(* Logix 5000 project; controller TFF vendor 1 type 14 code 107 rev 33.11; software revision 33.04; part 15 of 38 *)
(* tags used below, declared in another part *)
   ActionCode : DINT;   // Action Code
   AutoRunTimer : TIMER;   // Auto Run Timer
   Clear : BOOL;   // Clear Operation Table Flag
   Criteria1Code : DINT;   // Criteria 1 Code
   Criteria2Code : DINT;   // Criteria 2 Code
   CriteriaMet : BOOL;   // Criteria Met
   DownloadONS : BOOL;
   ErrorCheck : BOOL;   // Error Check Flag
   PhaseClear : BOOL;   // Phase Clear
   PhaseNumber : DINT;   // Phase FOR NEXT Index
   PreRunLog : BOOL;   // Log Pre Run Set Points
   Run : BOOL;   // Operation Run Status
   RunONS : BOOL;   // Run Command One-Shot
   Structure : DINT;   // Structure code
   Value : REAL;   // Temp Value
   AlarmControl : AlarmControl;   // Alarm Control
   CCPSystem : CCPSystem;   // CCP System Data
   CPU_Scanning : BOOL;   // System Scanning Flag
   Memory_Data : Memory_Data;
   Memory_Message : MESSAGE;   // Data for Message instruction read Memory informations
   Memory_Temp : INT[29];   // Destination elements for message read Memory informations
   Operation : Operation[6,251];   // Operation Table
   PCDateTime : DINT[7];   // Date/Time Array from PC
   Phase : Phases[6];   // Phase Control Array
   Phase0 : ALIAS FOR Phase[0];   // Phase 0
   PLCFault : FaultRecordType;   // PLC Major Fault Record
   Prompt : Prompt[7];   // Prompt Array
   Prompt0 : ALIAS FOR Prompt[0];   // Phase 0 Prompt
   Prompt1 : ALIAS FOR Prompt[1];   // Phase 1 Prompt
   Prompt2 : ALIAS FOR Prompt[2];   // Phase 2 Prompt
   Prompt3 : ALIAS FOR Prompt[3];   // Phase 3 Prompt
   Prompt4 : ALIAS FOR Prompt[4];   // Phase 4 Prompt
   Prompt5 : ALIAS FOR Prompt[5];   // Phase 5 Prompt
   ResumeDownloadFromHOLD : BOOL;   // Resume Download From HOLD
   TimerControl : TimerControl;   // Timer Control
   Timers : Timers[22];   // Timer Array
   YA10 : ALIAS FOR DigitalPoint[59];
(* CCPSystem, continued *)

ROUTINE Prompt   (* ladder *)
// Operator Prompt Routine
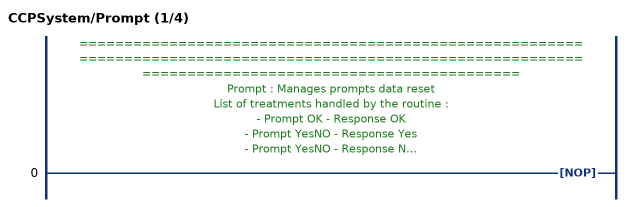
   // ==========================================================================================================================================================
   //                                                                                                                       Prompt : Manages prompts data reset
   //                                                     List of treatments handled by the routine :
   //                                                          - Prompt OK - Response OK
   //                                                          - Prompt YesNO - Response Yes
   //                                                          - Prompt YesNO - Response No
   //                                                     -----------------------------------------------------------------------------------------------------------------------------------------------------
   //                                                     History
   // 		2019-DEC-24 - Merck - Q. Spindler - Initial version for Candidate Release 1.00.00.00.a
   // 		2022-SEP-20 - Actemium - J. Jaekel - Modification for Candidate Release 1.01.00.01.a
   // - Add condition to avoid discarding the prompt response on other phases than 0
   // ============================================================================================================================
   // ============================
   0: NOP();
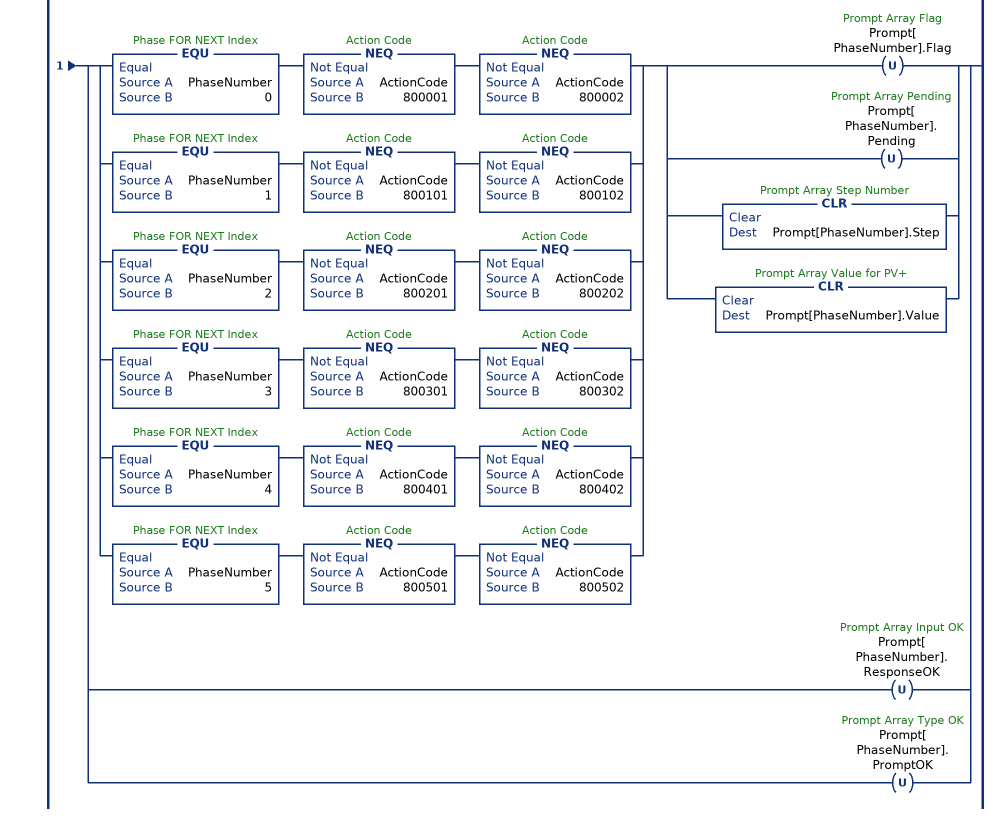
   // Prompt OK - Response OK
   // ==========================================================================================================================================================
   1: XIC(Prompt[PhaseNumber].PromptOK)XIC(Prompt[PhaseNumber].ResponseOK)[XIC(CriteriaMet) ,XIC(Phase[PhaseNumber].JumpPLC) ,EQU(PhaseNumber,0) NEQ(Criteria1Code,800003) NEQ(Criteria2Code,800003) ,EQU(PhaseNumber,1) NEQ(Criteria1Code,800103) NEQ(Criteria2Code,800103) ,EQU(PhaseNumber,2) NEQ(Criteria1Code,800203) NEQ(Criteria2Code,800203) ,EQU(PhaseNumber,3) NEQ(Criteria1Code,800303) NEQ(Criteria2Code,800303) ,EQU(PhaseNumber,4) NEQ(Criteria1Code,800403) NEQ(Criteria2Code,800403) ,EQU(PhaseNumber,5) NEQ(Criteria1Code,800503) NEQ(Criteria2Code,800503) ][[EQU(PhaseNumber,0) NEQ(ActionCode,800001) NEQ(ActionCode,800002) ,EQU(PhaseNumber,1) NEQ(ActionCode,800101) NEQ(ActionCode,800102) ,EQU(PhaseNumber,2) NEQ(ActionCode,800201) NEQ(ActionCode,800202) ,EQU(PhaseNumber,3) NEQ(ActionCode,800301) NEQ(ActionCode,800302) ,EQU(PhaseNumber,4) NEQ(ActionCode,800401) NEQ(ActionCode,800402) ,EQU(PhaseNumber,5) NEQ(ActionCode,800501) NEQ(ActionCode,800502) ] [OTU(Prompt[PhaseNumber].Flag) ,OTU(Prompt[PhaseNumber].Pending) ,CLR(Prompt[PhaseNumber].Step) ,CLR(Prompt[PhaseNumber].Value) ] ,OTU(Prompt[PhaseNumber].ResponseOK) ,OTU(Prompt[PhaseNumber].PromptOK) ];
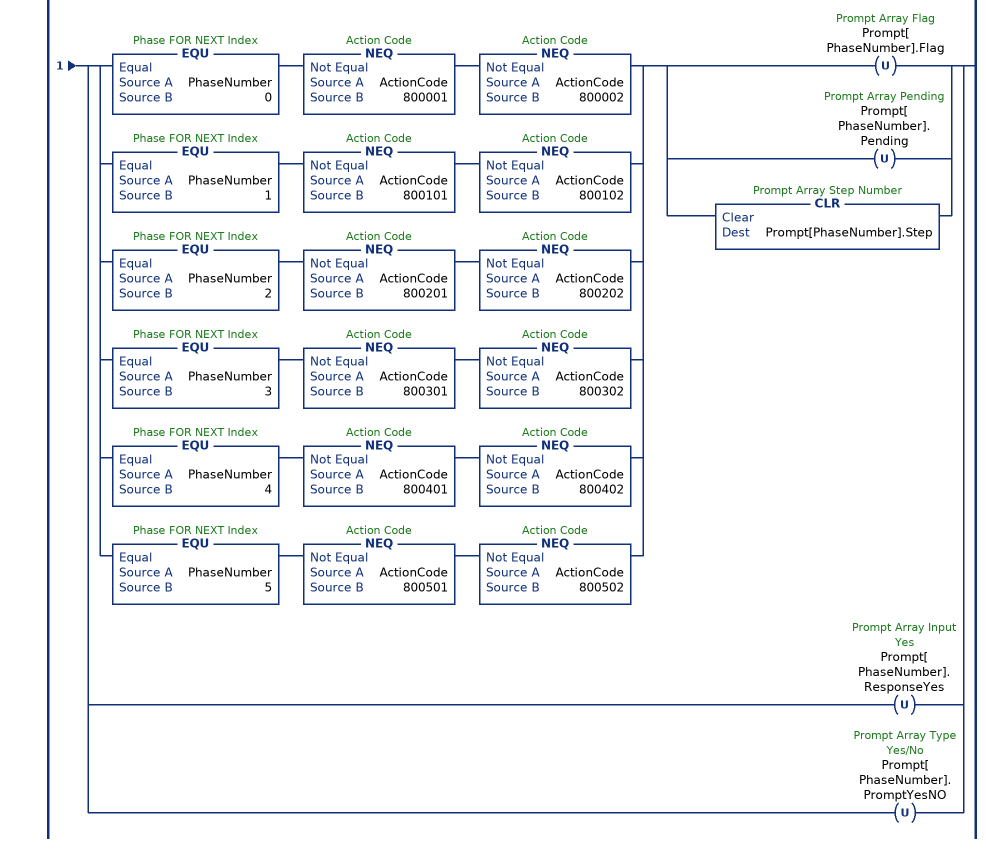
   // Prompt YesNO - Response Yes
   // ==========================================================================================================================================================
   2: XIC(Prompt[PhaseNumber].PromptYesNO)XIC(Prompt[PhaseNumber].ResponseYes)[XIC(CriteriaMet) ,XIC(Phase[PhaseNumber].JumpPLC) ,EQU(PhaseNumber,0) NEQ(Criteria1Code,800004) NEQ(Criteria2Code,800004) ,EQU(PhaseNumber,1) NEQ(Criteria1Code,800104) NEQ(Criteria2Code,800104) ,EQU(PhaseNumber,2) NEQ(Criteria1Code,800204) NEQ(Criteria2Code,800204) ,EQU(PhaseNumber,3) NEQ(Criteria1Code,800304) NEQ(Criteria2Code,800304) ,EQU(PhaseNumber,4) NEQ(Criteria1Code,800404) NEQ(Criteria2Code,800404) ,EQU(PhaseNumber,5) NEQ(Criteria1Code,800504) NEQ(Criteria2Code,800504) ][[EQU(PhaseNumber,0) NEQ(ActionCode,800001) NEQ(ActionCode,800002) ,EQU(PhaseNumber,1) NEQ(ActionCode,800101) NEQ(ActionCode,800102) ,EQU(PhaseNumber,2) NEQ(ActionCode,800201) NEQ(ActionCode,800202) ,EQU(PhaseNumber,3) NEQ(ActionCode,800301) NEQ(ActionCode,800302) ,EQU(PhaseNumber,4) NEQ(ActionCode,800401) NEQ(ActionCode,800402) ,EQU(PhaseNumber,5) NEQ(ActionCode,800501) NEQ(ActionCode,800502) ] [OTU(Prompt[PhaseNumber].Flag) ,OTU(Prompt[PhaseNumber].Pending) ,CLR(Prompt[PhaseNumber].Step) ] ,OTU(Prompt[PhaseNumber].ResponseYes) ,OTU(Prompt[PhaseNumber].PromptYesNO) ];
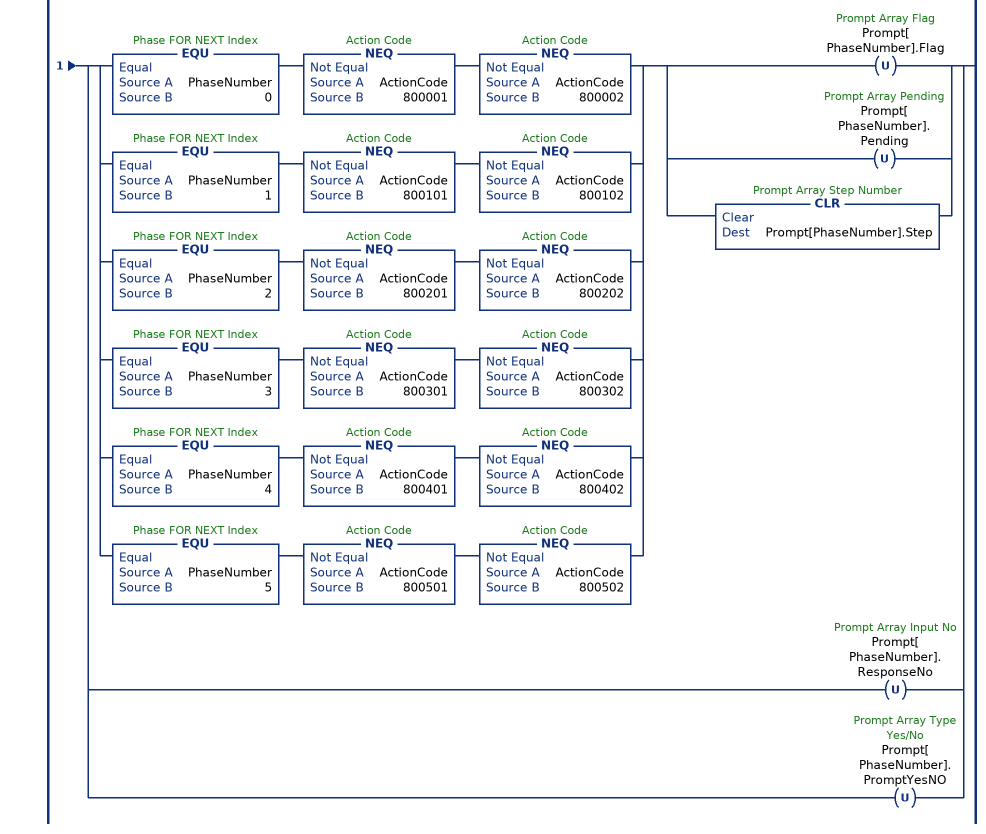
   // Prompt YesNO - Response No
   // ==========================================================================================================================================================
   3: XIC(Prompt[PhaseNumber].PromptYesNO)XIC(Prompt[PhaseNumber].ResponseNo)[XIC(CriteriaMet) ,XIC(Phase[PhaseNumber].JumpPLC) ,EQU(PhaseNumber,0) NEQ(Criteria1Code,800005) NEQ(Criteria2Code,800005) ,EQU(PhaseNumber,1) NEQ(Criteria1Code,800105) NEQ(Criteria2Code,800105) ,EQU(PhaseNumber,2) NEQ(Criteria1Code,800205) NEQ(Criteria2Code,800205) ,EQU(PhaseNumber,3) NEQ(Criteria1Code,800305) NEQ(Criteria2Code,800305) ,EQU(PhaseNumber,4) NEQ(Criteria1Code,800405) NEQ(Criteria2Code,800405) ,EQU(PhaseNumber,5) NEQ(Criteria1Code,800505) NEQ(Criteria2Code,800505) ][[EQU(PhaseNumber,0) NEQ(ActionCode,800001) NEQ(ActionCode,800002) ,EQU(PhaseNumber,1) NEQ(ActionCode,800101) NEQ(ActionCode,800102) ,EQU(PhaseNumber,2) NEQ(ActionCode,800201) NEQ(ActionCode,800202) ,EQU(PhaseNumber,3) NEQ(ActionCode,800301) NEQ(ActionCode,800302) ,EQU(PhaseNumber,4) NEQ(ActionCode,800401) NEQ(ActionCode,800402) ,EQU(PhaseNumber,5) NEQ(ActionCode,800501) NEQ(ActionCode,800502) ] [OTU(Prompt[PhaseNumber].Flag) ,OTU(Prompt[PhaseNumber].Pending) ,CLR(Prompt[PhaseNumber].Step) ] ,OTU(Prompt[PhaseNumber].ResponseNo) ,OTU(Prompt[PhaseNumber].PromptYesNO) ];
END_ROUTINE

ROUTINE Start   (* ladder *)
// Operation Start Routine
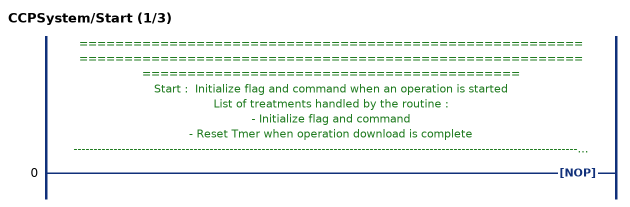
   // ==========================================================================================================================================================
   //                                                                                                      Start :  Initialize flag and command when an operation is started
   //                                                     List of treatments handled by the routine :
   //                                                          - Initialize flag and command
   //                                                          - Reset Tmer when operation download is complete
   //                                                     -----------------------------------------------------------------------------------------------------------------------------------------------------
   //                                                     History
   // 		2019-DEC-24 - Merck - Q. Spindler - Initial version for Candidate Release 1.00.00.00.a
   // ========================================================================================================================================================
   0: NOP();
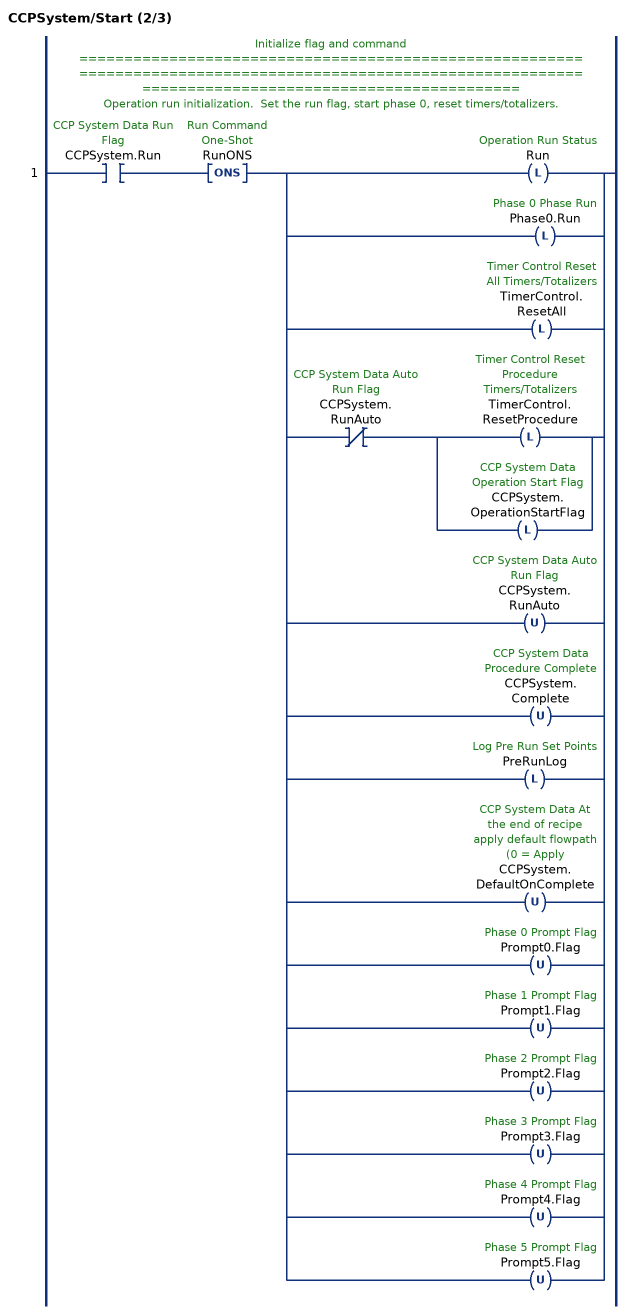
   // Initialize flag and command
   // ==========================================================================================================================================================
   // Operation run initialization.  Set the run flag, start phase 0, reset timers/totalizers.
   1: XIC(CCPSystem.Run)ONS(RunONS)[OTL(Run) ,OTL(Phase0.Run) ,OTL(TimerControl.ResetAll) ,XIO(CCPSystem.RunAuto) [OTL(TimerControl.ResetProcedure) ,OTL(CCPSystem.OperationStartFlag) ] ,OTU(CCPSystem.RunAuto) ,OTU(CCPSystem.Complete) ,OTL(PreRunLog) ,OTU(CCPSystem.DefaultOnComplete) ,OTU(Prompt0.Flag) ,OTU(Prompt1.Flag) ,OTU(Prompt2.Flag) ,OTU(Prompt3.Flag) ,OTU(Prompt4.Flag) ,OTU(Prompt5.Flag) ];
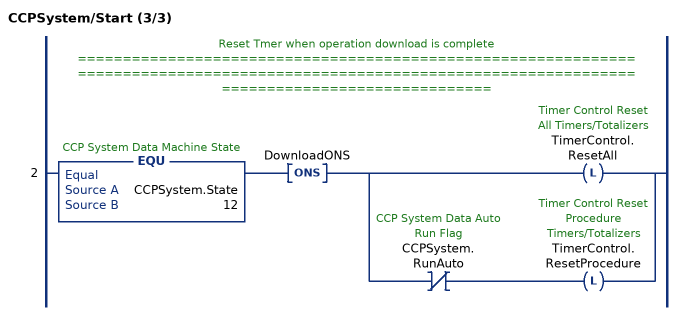
   // Reset Tmer when operation download is complete
   // ==========================================================================================================================================================
   2: EQU(CCPSystem.State,12)ONS(DownloadONS)[OTL(TimerControl.ResetAll) ,XIO(CCPSystem.RunAuto) OTL(TimerControl.ResetProcedure) ];
END_ROUTINE

ROUTINE State   (* ladder *)
// Machine State Routine
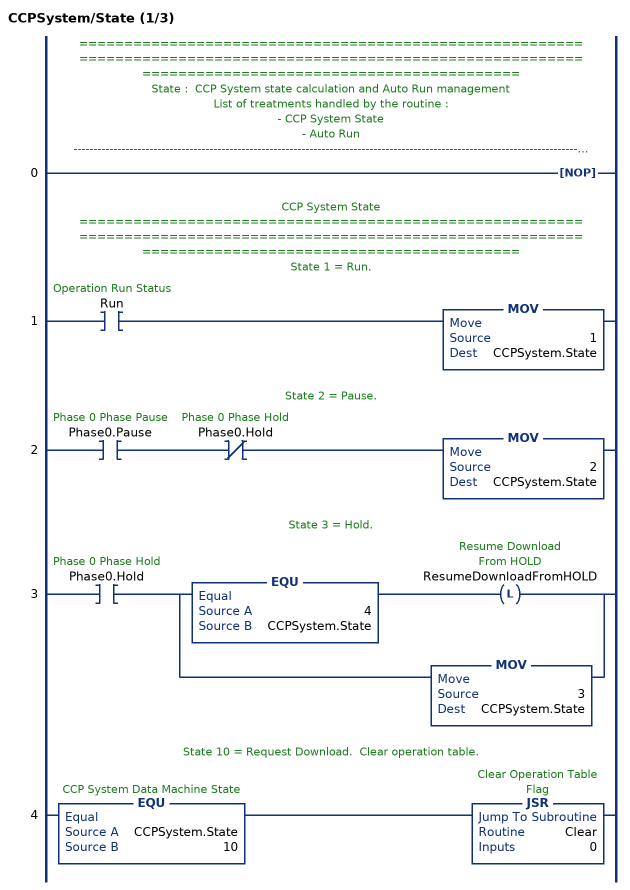
   // ==========================================================================================================================================================
   //                                                                                                  State :  CCP System state calculation and Auto Run management
   //                                                     List of treatments handled by the routine :
   //                                                          - CCP System State
   //                                                          - Auto Run
   //                                                     -----------------------------------------------------------------------------------------------------------------------------------------------------
   //                                                     History
   // 		2019-DEC-24 - Merck - Q. Spindler - Initial version for Candidate Release 1.00.00.00.a
   // 		2021-APR-22 - Merck - Q. Spindler - Modifications for Candidate Release 1.00.00.00.e
   // - Add of Resume Download From HOLD state
   // ========================================================================================================================================================
   0: NOP();
   // CCP System State
   // ==========================================================================================================================================================
   // State 1 = Run.
   1: XIC(Run)MOV(1,CCPSystem.State);
   // State 2 = Pause.
   2: XIC(Phase0.Pause)XIO(Phase0.Hold)MOV(2,CCPSystem.State);
   // State 3 = Hold.
   3: XIC(Phase0.Hold)[EQU(4,CCPSystem.State) OTL(ResumeDownloadFromHOLD) ,MOV(3,CCPSystem.State) ];
   // State 10 = Request Download.  Clear operation table.
   4: EQU(CCPSystem.State,10)JSR(Clear,0);
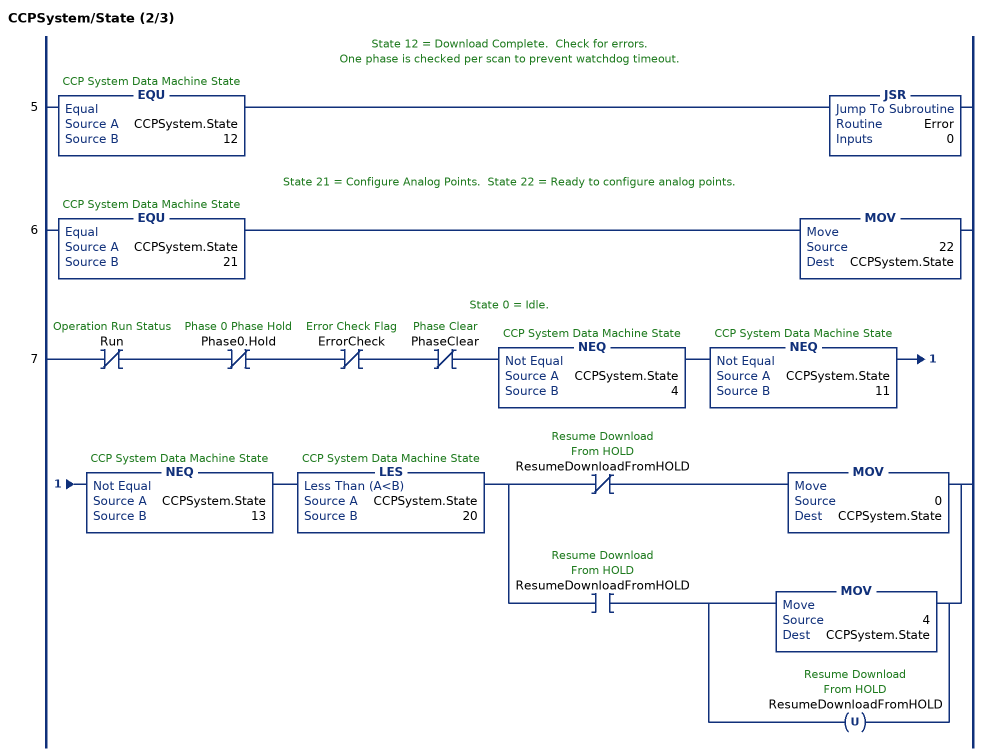
   // State 12 = Download Complete.  Check for errors.
   // One phase is checked per scan to prevent watchdog timeout.
   5: EQU(CCPSystem.State,12)JSR(Error,0);
   // State 21 = Configure Analog Points.  State 22 = Ready to configure analog points.
   6: EQU(CCPSystem.State,21)MOV(22,CCPSystem.State);
   // State 0 = Idle.
   7: XIO(Run)XIO(Phase0.Hold)XIO(ErrorCheck)XIO(PhaseClear)NEQ(CCPSystem.State,4)NEQ(CCPSystem.State,11)NEQ(CCPSystem.State,13)LES(CCPSystem.State,20)[XIO(ResumeDownloadFromHOLD) MOV(0,CCPSystem.State) ,XIC(ResumeDownloadFromHOLD) [MOV(4,CCPSystem.State) ,OTU(ResumeDownloadFromHOLD) ] ];
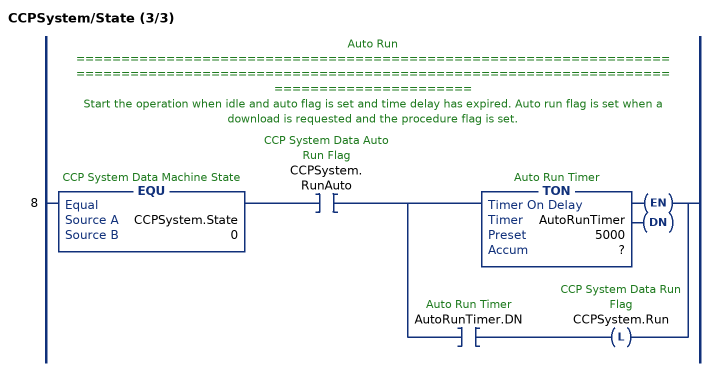
   // Auto Run
   // ==========================================================================================================================================================
   // Start the operation when idle and auto flag is set and time delay has expired. Auto run flag is set when a download is requested and the procedure flag is set.
   8: EQU(CCPSystem.State,0)XIC(CCPSystem.RunAuto)[TON(AutoRunTimer,?,?) ,XIC(AutoRunTimer.DN) OTL(CCPSystem.Run) ];
END_ROUTINE
END_PROGRAM

PROGRAM ControllerFaultRoutine   (* main routine FaultRoutine *)

ROUTINE FaultRoutine   (* ladder *)
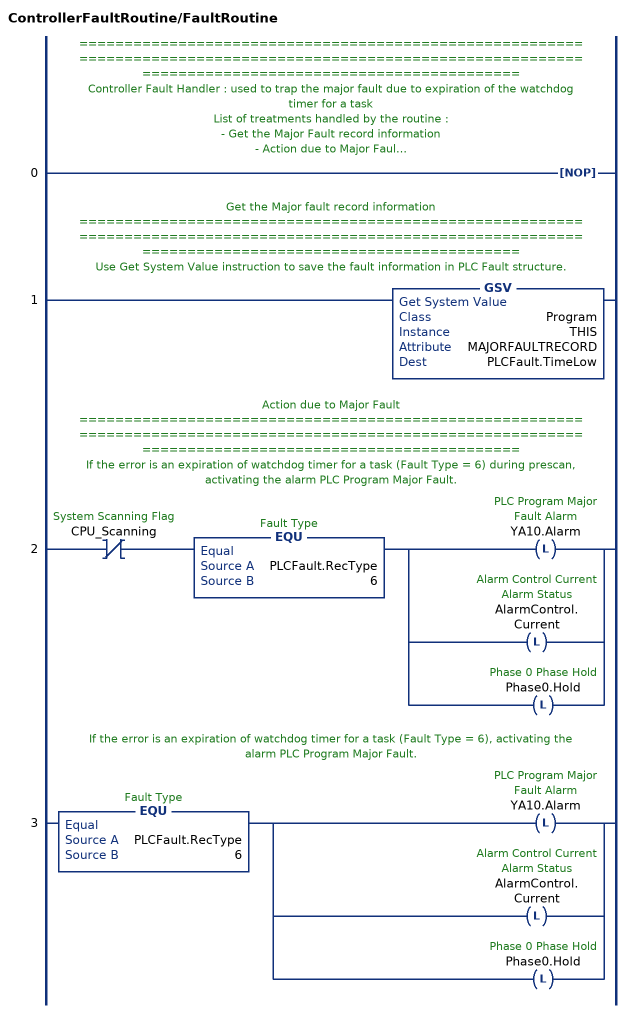
   // ==========================================================================================================================================================
   //                                                                                 Controller Fault Handler : used to trap the major fault due to expiration of the watchdog timer for a task
   //                                                     List of treatments handled by the routine :
   //                                                          - Get the Major Fault record information
   //                                                          - Action due to Major Fault
   //                                                     -----------------------------------------------------------------------------------------------------------------------------------------------------
   //                                                     History
   // 		2019-DEC-24 - Merck - Q. Spindler - Initial version for Candidate Release 1.00.00.00.a
   // ==========================================================================================================================================================
   0: NOP();
   // Get the Major fault record information
   // ==========================================================================================================================================================
   // Use Get System Value instruction to save the fault information in PLC Fault structure.
   1: GSV(Program,THIS,MAJORFAULTRECORD,PLCFault.TimeLow);
   // Action due to Major Fault
   // ==========================================================================================================================================================
   // If the error is an expiration of watchdog timer for a task (Fault Type = 6) during prescan, activating the alarm PLC Program Major Fault.
   2: XIO(CPU_Scanning)EQU(PLCFault.RecType,6)[OTL(YA10.Alarm) ,OTL(AlarmControl.Current) ,OTL(Phase0.Hold) ];
   // If the error is an expiration of watchdog timer for a task (Fault Type = 6), activating the alarm PLC Program Major Fault.
   3: EQU(PLCFault.RecType,6)[OTL(YA10.Alarm) ,OTL(AlarmControl.Current) ,OTL(Phase0.Hold) ];
END_ROUTINE
END_PROGRAM

PROGRAM MainProgram   (* main routine MainRoutine, fault routine FaultRoutine *)
// Date/Time Synchronization
VAR
   Address : DINT := 9;   // Temp Address used in Time Loop
   AddressTotalizer : DINT := 20;   // Temp Address used in modPhaseTotal
   Index : DINT := 2;   // Index
   PLCDST : SINT;   // Current PLC Day Light Saving
   PLCTimeZoneString : STRING := 'UTC+00:00 Coordinated Universal Time';   // Current PLC TimeZone
   SCL : SCALE := (In := -4.0, InRawMax := 99999.0, InEUMax := 999.99, Out := -0.04, MinAlarm := 1);
   TimeZoneUTC0 : STRING := 'UTC+00:00 Coordinated Universal Time';   // String value for Time zone UTC 0
END_VAR

ROUTINE FaultRoutine   (* ladder *)
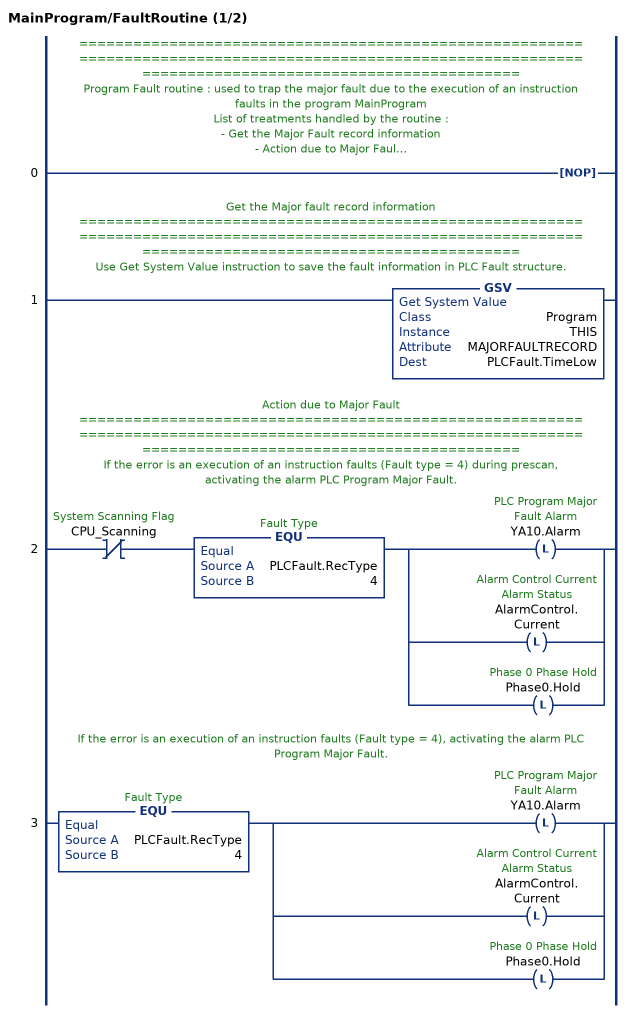
   // ==========================================================================================================================================================
   //                                                               Program Fault routine : used to trap the major fault due to the execution of an instruction faults in the program MainProgram
   //                                                     List of treatments handled by the routine :
   //                                                          - Get the Major Fault record information
   //                                                          - Action due to Major Fault
   //                                                     -----------------------------------------------------------------------------------------------------------------------------------------------------
   //                                                     History
   // 		2019-DEC-24 - Merck - Q. Spindler - Initial version for Candidate Release 1.00.00.00.a
   // ==========================================================================================================================================================
   0: NOP();
   // Get the Major fault record information
   // ==========================================================================================================================================================
   // Use Get System Value instruction to save the fault information in PLC Fault structure.
   1: GSV(Program,THIS,MAJORFAULTRECORD,PLCFault.TimeLow);
   // Action due to Major Fault
   // ==========================================================================================================================================================
   // If the error is an execution of an instruction faults (Fault type = 4) during prescan, activating the alarm PLC Program Major Fault.
   2: XIO(CPU_Scanning)EQU(PLCFault.RecType,4)[OTL(YA10.Alarm) ,OTL(AlarmControl.Current) ,OTL(Phase0.Hold) ];
   // If the error is an execution of an instruction faults (Fault type = 4), activating the alarm PLC Program Major Fault.
   3: EQU(PLCFault.RecType,4)[OTL(YA10.Alarm) ,OTL(AlarmControl.Current) ,OTL(Phase0.Hold) ];
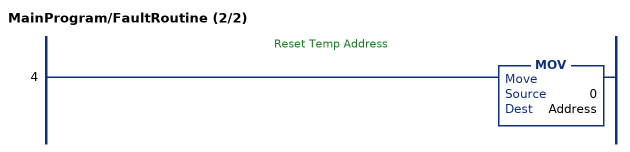
   // Reset Temp Address
   4: MOV(0,Address);
END_ROUTINE

ROUTINE MainRoutine   (* ladder *)
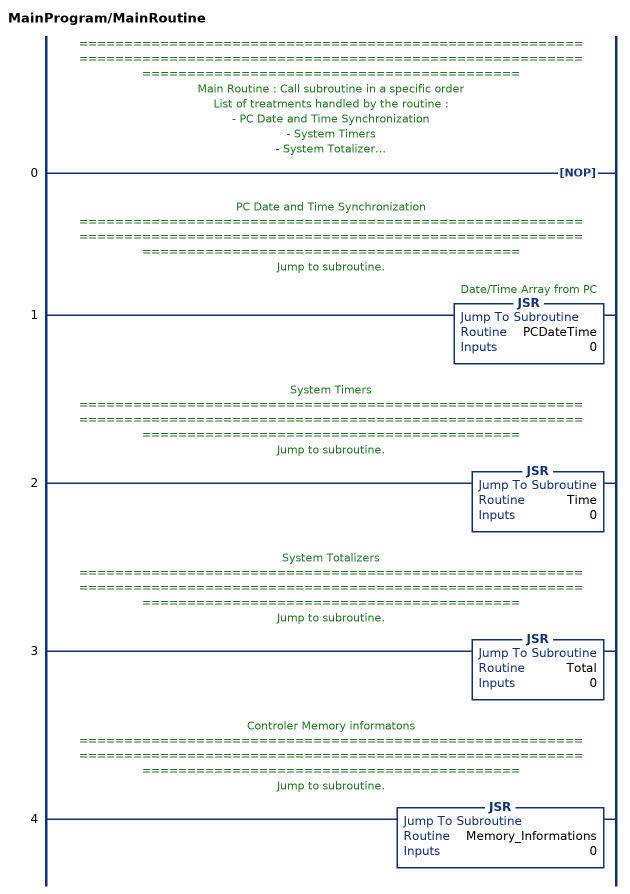
   // ==========================================================================================================================================================
   //                                                                                                            Main Routine : Call subroutine in a specific order
   //                                                     List of treatments handled by the routine :
   //                                                          - PC Date and Time Synchronization
   //                                                          - System Timers
   //                                                          - System Totalizers
   //                                                           - Controler Memory informatons
   //                                                     -----------------------------------------------------------------------------------------------------------------------------------------------------
   //                                                     History
   // 		2019-DEC-24 - Merck - Q. Spindler - Initial version for Candidate Release 1.00.00.00.a
   // 		2021-NOV-17 - Merck - Q.Spindler - Modifications for Candidate Release 1.01.00.00.a
   // - Add Memory_Information Call
   // ==========================================================================================================================================================
   0: NOP();
   // PC Date and Time Synchronization
   // ==========================================================================================================================================================
   // Jump to subroutine.
   1: JSR(PCDateTime,0);
   // System Timers
   // ==========================================================================================================================================================
   // Jump to subroutine.
   2: JSR(Time,0);
   // System Totalizers
   // ==========================================================================================================================================================
   // Jump to subroutine.
   3: JSR(Total,0);
   // Controler Memory informatons
   // ==========================================================================================================================================================
   // Jump to subroutine.
   4: JSR(Memory_Informations,0);
END_ROUTINE

ROUTINE Memory_Data   (* ladder *)
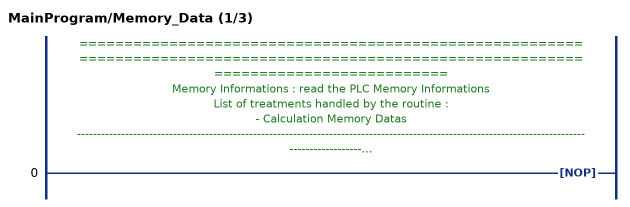
   // ==========================================================================================================================================
   // Memory Informations : read the PLC Memory Informations
   // List of treatments handled by the routine :
   // - Calculation Memory Datas
   //                                                     --------------------------------------------------------------------------------------------------------------------------------------------------
   // History
   // 		2021-Nov-17 - Merck - Q.Spindler - Initial version for Candidate Release 1.01.00.00.a
   // ==========================================================================================================================================
   0: NOP();
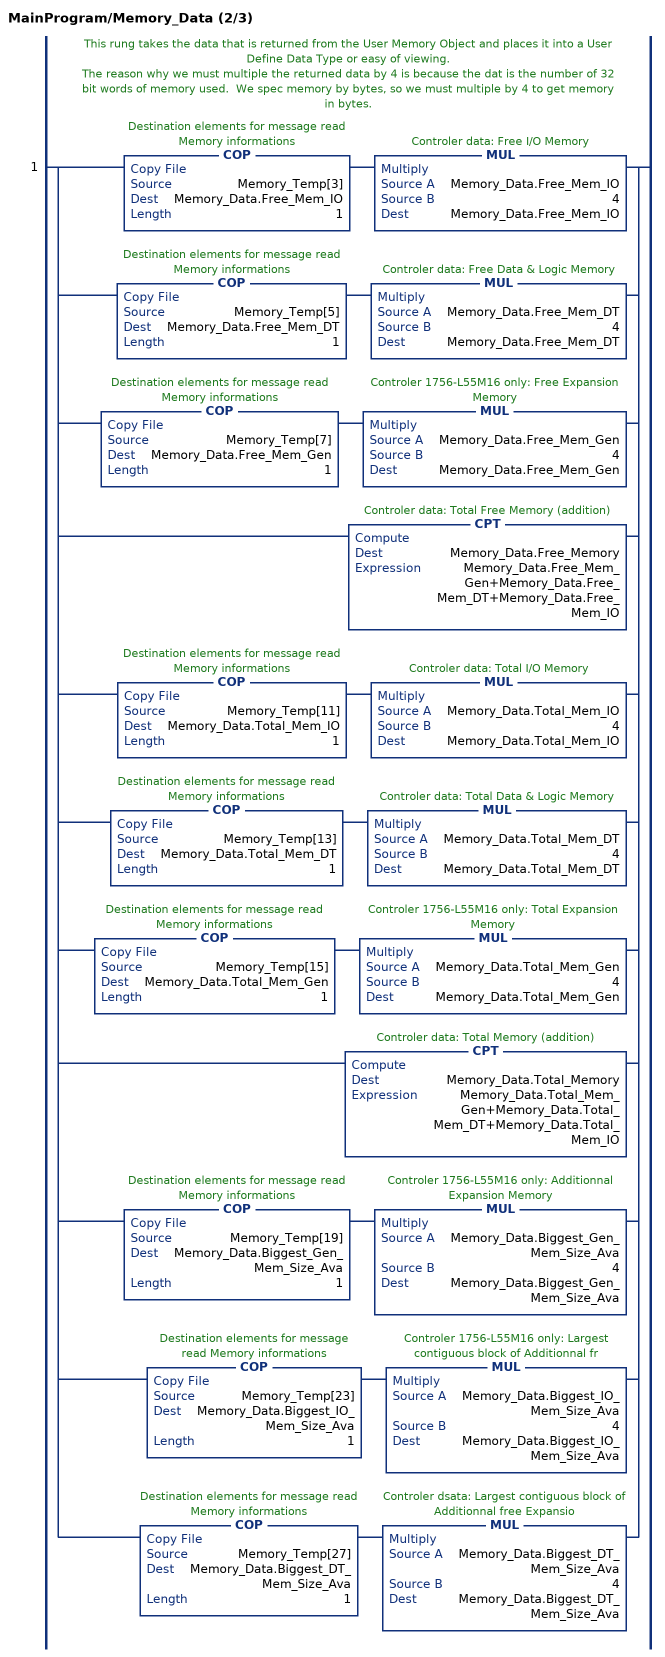
   // This rung takes the data that is returned from the User Memory Object and places it into a User Define Data Type or easy of viewing.
   // The reason why we must multiple the returned data by 4 is because the dat is the number of 32 bit words of memory used.  We spec memory by bytes, so we must multiple by 4 to get memory in bytes.
   1: [COP(Memory_Temp[3],Memory_Data.Free_Mem_IO,1) MUL(Memory_Data.Free_Mem_IO,4,Memory_Data.Free_Mem_IO) ,COP(Memory_Temp[5],Memory_Data.Free_Mem_DT,1) MUL(Memory_Data.Free_Mem_DT,4,Memory_Data.Free_Mem_DT) ,COP(Memory_Temp[7],Memory_Data.Free_Mem_Gen,1) MUL(Memory_Data.Free_Mem_Gen,4,Memory_Data.Free_Mem_Gen) ,CPT(Memory_Data.Free_Memory,Memory_Data.Free_Mem_Gen+Memory_Data.Free_Mem_DT+Memory_Data.Free_Mem_IO) ,COP(Memory_Temp[11],Memory_Data.Total_Mem_IO,1) MUL(Memory_Data.Total_Mem_IO,4,Memory_Data.Total_Mem_IO) ,COP(Memory_Temp[13],Memory_Data.Total_Mem_DT,1) MUL(Memory_Data.Total_Mem_DT,4,Memory_Data.Total_Mem_DT) ,COP(Memory_Temp[15],Memory_Data.Total_Mem_Gen,1) MUL(Memory_Data.Total_Mem_Gen,4,Memory_Data.Total_Mem_Gen) ,CPT(Memory_Data.Total_Memory,Memory_Data.Total_Mem_Gen+Memory_Data.Total_Mem_DT+Memory_Data.Total_Mem_IO) ,COP(Memory_Temp[19],Memory_Data.Biggest_Gen_Mem_Size_Ava,1) MUL(Memory_Data.Biggest_Gen_Mem_Size_Ava,4,Memory_Data.Biggest_Gen_Mem_Size_Ava) ,COP(Memory_Temp[23],Memory_Data.Biggest_IO_Mem_Size_Ava,1) MUL(Memory_Data.Biggest_IO_Mem_Size_Ava,4,Memory_Data.Biggest_IO_Mem_Size_Ava) ,COP(Memory_Temp[27],Memory_Data.Biggest_DT_Mem_Size_Ava,1) MUL(Memory_Data.Biggest_DT_Mem_Size_Ava,4,Memory_Data.Biggest_DT_Mem_Size_Ava) ];
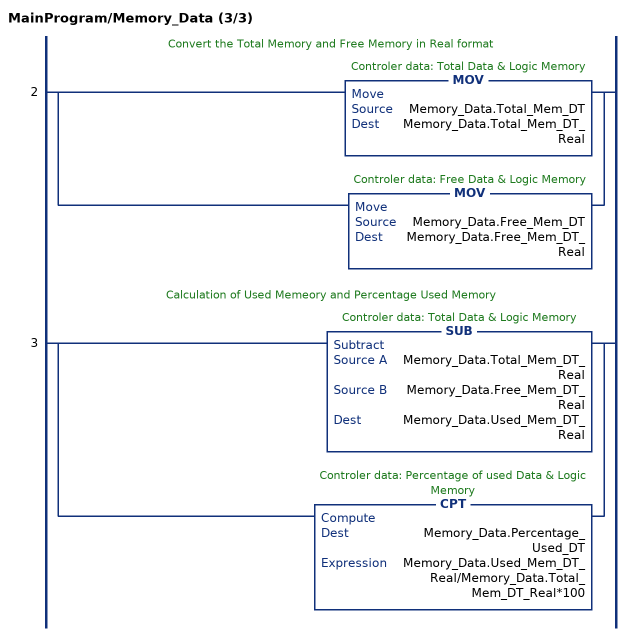
   // Convert the Total Memory and Free Memory in Real format
   2: [MOV(Memory_Data.Total_Mem_DT,Memory_Data.Total_Mem_DT_Real) ,MOV(Memory_Data.Free_Mem_DT,Memory_Data.Free_Mem_DT_Real) ];
   // Calculation of Used Memeory and Percentage Used Memory
   3: [SUB(Memory_Data.Total_Mem_DT_Real,Memory_Data.Free_Mem_DT_Real,Memory_Data.Used_Mem_DT_Real) ,CPT(Memory_Data.Percentage_Used_DT,Memory_Data.Used_Mem_DT_Real/Memory_Data.Total_Mem_DT_Real*100) ];
END_ROUTINE

ROUTINE Memory_Informations   (* ladder *)
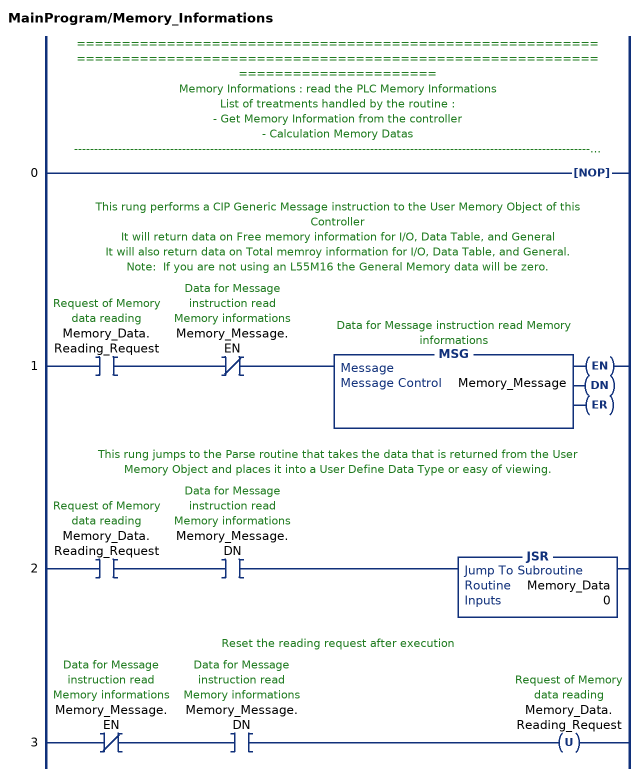
   // ==========================================================================================================================================
   // Memory Informations : read the PLC Memory Informations
   // List of treatments handled by the routine :
   // - Get Memory Information from the controller
   // - Calculation Memory Datas
   //                                                     --------------------------------------------------------------------------------------------------------------------------------------------------
   // History
   // 		2021-Nov-17 - Merck - Q.Spindler - Initial version for Candidate Release 1.01.00.00.a
   // ==========================================================================================================================================
   0: NOP();
   // This rung performs a CIP Generic Message instruction to the User Memory Object of this Controller
   // It will return data on Free memory information for I/O, Data Table, and General
   // It will also return data on Total memroy information for I/O, Data Table, and General.
   // Note:  If you are not using an L55M16 the General Memory data will be zero.
   1: XIC(Memory_Data.Reading_Request)XIO(Memory_Message.EN)MSG(Memory_Message);
   // This rung jumps to the Parse routine that takes the data that is returned from the User Memory Object and places it into a User Define Data Type or easy of viewing.
   2: XIC(Memory_Data.Reading_Request)XIC(Memory_Message.DN)JSR(Memory_Data,0);
   // Reset the reading request after execution
   3: XIO(Memory_Message.EN)XIC(Memory_Message.DN)OTU(Memory_Data.Reading_Request);
END_ROUTINE
